// TIA Portal V20 export
TYPE "Wartungszähler_Weg"
   STRUCT
      Gesamtweg : DInt;
      Weg_soll : DInt;
      Weg_seit_Wartung : DInt;
      Weg_bis_Wartung : DInt;
      Zähler_reset : Bool;
      SM_Wartung_fällig : Bool;
   END_STRUCT;
END_TYPE
